(* IEC 61131-3 sources: Test-Git_ESME26/00_Initial Project_LB.fbsproj/M660.device.xml.v3^/Plc Logic.plclogic.xml.v3^/Application.application.xml.v3^/Application, 1 file *)

(* ---- SR_Application.prg.st ---- *)
PROGRAM SR_Application
VAR
	fbLogicEnc : MOIN.FB_LogicalEncoder;
	fbVirtualMaster : MOIN.FB_ControlledAxis;

	xTest		: BOOL;
END_VAR

xTest := FALSE;
//GitHub test
//questo testo appare solo nella parte del Branch
